Fanuc KAREL source: KA00174.KL

PROGRAM KA00174
%NOLOCKGROUP
VAR
  SRC: ARRAY[4] OF STRING[20]
  DST: ARRAY[4] OF BOOLEAN
BEGIN
  DST = SRC
END KA00174
